SUBAPPLICATION AR_TO_Q_Publish_Fast_OPC (* AR-Wert per OPC-UA ungedrosselt publizieren (Regelung), VT-Anzeige auf max. 1 Update/500 ms gedrosselt *)
  (* Standard: 61499-2; Description: Copyright (c) 2026 Meisterschulen am Ostbahnhof This program and the accompanying materials are made available under the terms of the Eclipse Public License 2.0 which is available at https://www.eclipse.org/legal/epl-2.0/ SPDX-License-Identifier: EPL-2.0 *)
  (* Version 1.0, 2026-10-30, Franz Höpfinger, Meisterschulen am Ostbahnhof, Kopie von AR_TO_Q_Publish_OPC (v1.2), RateLimit_Anzeige wieder HINTER den Split, nur vor Q_NumericValue: AR_PUBLISH (Self-Subscribe der Regelung, z.B. Fahrwerk_Mittelpunkt_Automatik) ungedrosselt. Franz: Regelung muss schnell sein, die Anzeige darf hinterherhinken. *)
  PACKAGE MyLib::sys;
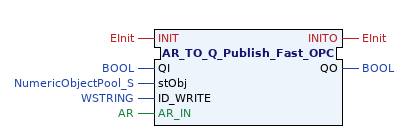
  EVENT_INPUT
    INIT : EInit; (* Initialization Request *)
  END_EVENT
  EVENT_OUTPUT
    INITO : EInit; (* Initialization Confirm *)
  END_EVENT
  VAR_INPUT
    QI : BOOL := TRUE; (* Quality Input - TRUE to enable service *)
    stObj : logiBUS::utils::conversion::phys::NumericObjectPool_S; (* Object pool properties der VT-Zahlenvariable (u16ObjId, scale, offset, decimals) - z.B. FBs::const::DefaultPool_Numeric::NumberVariable_X_N *)
    ID_WRITE : WSTRING; (* Publish-Adresse (REAL, ACTION=PUBLISH), lokal oder stationsuebergreifend *)
  END_VAR
  VAR_OUTPUT
    QO : BOOL; (* Quality Output - TRUE if service executed successfully *)
  END_VAR
  SOCKETS
    AR_IN : adapter::types::unidirectional::AR; (* Physikalischer Wert (bereits skaliert) *)
  END_SOCKETS
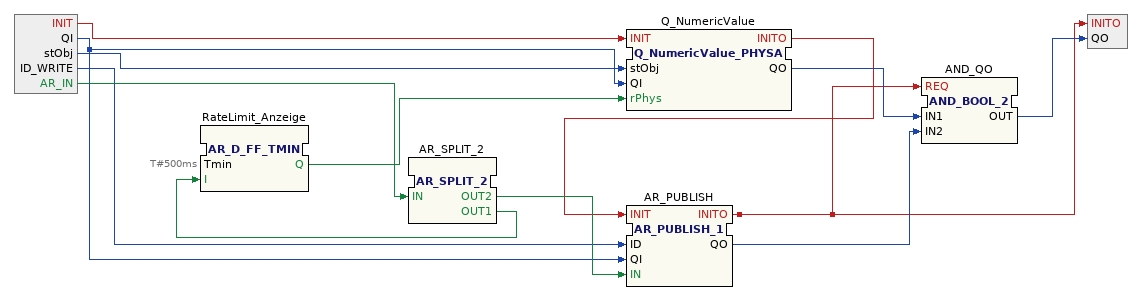
  FBS
    AR_SPLIT_2 : adapter::events::unidirectional::AR_SPLIT_2;
    RateLimit_Anzeige : adapter::events::unidirectional::AR_D_FF_TMIN(Tmin := T#500ms); (* Drosselt nur die VT-Anzeige, AR_PUBLISH bleibt ungedrosselt *)
    Q_NumericValue : isobus::UT::Q::Q_NumericValue_PHYSA;
    AR_PUBLISH : adapter::net::AR_PUBLISH_1;
    AND_QO : iec61131::booleanOperators::AND_BOOL_2;
  END_FBS
  EVENT_CONNECTIONS
    INIT TO Q_NumericValue.INIT;
    Q_NumericValue.INITO TO AR_PUBLISH.INIT;
    AR_PUBLISH.INITO TO INITO;
    AR_PUBLISH.INITO TO AND_QO.REQ;
  END_CONNECTIONS
  DATA_CONNECTIONS
    stObj TO Q_NumericValue.stObj;
    ID_WRITE TO AR_PUBLISH.ID;
    QI TO Q_NumericValue.QI;
    QI TO AR_PUBLISH.QI;
    Q_NumericValue.QO TO AND_QO.IN1;
    AR_PUBLISH.QO TO AND_QO.IN2;
    AND_QO.OUT TO QO;
  END_CONNECTIONS
  ADAPTER_CONNECTIONS
    AR_IN TO AR_SPLIT_2.IN;
    AR_SPLIT_2.OUT2 TO AR_PUBLISH.IN;
    AR_SPLIT_2.OUT1 TO RateLimit_Anzeige.I;
    RateLimit_Anzeige.Q TO Q_NumericValue.rPhys;
  END_CONNECTIONS
END_SUBAPPLICATION
